(* IEC 61131-3 sources: volt/packages/volt-lsp-iec/libraries/Standard/3.5.18.0, 22 files *)

(* ---- CONCAT.pou ---- *)
FUNCTION CONCAT : STRING(255)
VAR_INPUT
	STR1 : STRING(255);
	STR2 : STRING(255);
END_VAR
VAR
	i : DINT;
	n : DINT;
END_VAR
(* STR2 after STR1, cut at the 255 the result holds *)
CONCAT := STR1;
n := UINT_TO_DINT(LEN_INTERNAL(STR1));
WHILE n + i < 255 AND STR2[i] <> 0 DO
	CONCAT[n + i] := STR2[i];
	i := i + 1;
END_WHILE
CONCAT[n + i] := 0;
END_FUNCTION

(* ---- DELETE.pou ---- *)
FUNCTION DELETE : STRING(255)
VAR_INPUT
	STR : STRING(255);
	LEN : INT;
	POS : INT;
END_VAR
VAR
	i : DINT;
	k : DINT;
	n : DINT;
	first : DINT;
	start : DINT;
	count : DINT;
END_VAR
(* LEN characters from POS, counting from 1. POSITION 0 IS NOT "DO NOTHING": the range starts at POS - 1, which may
   be negative, and what goes is the part of [POS - 1, POS - 1 + LEN) inside the string. DELETE('abcde', 2, 0) is
   'bcde' (measured str_delete_at_zero, 2026-09-19). *)
DELETE := STR;
IF LEN > 0 THEN
	n := UINT_TO_DINT(LEN_INTERNAL(STR));
	first := INT_TO_DINT(POS) - 1;
	start := MAX(first, 0);
	count := INT_TO_DINT(LEN) + MIN(first, 0);
	IF count > 0 AND start < n THEN
		k := start;
		FOR i := MIN(start + count, n) TO n - 1 DO
			DELETE[k] := STR[i];
			k := k + 1;
		END_FOR
		DELETE[k] := 0;
	END_IF
END_IF
END_FUNCTION

(* ---- FIND.pou ---- *)
FUNCTION FIND : INT
VAR_INPUT
	STR1 : STRING(255);
	STR2 : STRING(255);
END_VAR
VAR
	i : DINT;
	j : DINT;
	n1 : DINT;
	n2 : DINT;
END_VAR
(* where STR2 first starts in STR1, counting from 1; 0 when it does not occur, and FIND of '' is 0 *)
n1 := UINT_TO_DINT(LEN_INTERNAL(STR1));
n2 := UINT_TO_DINT(LEN_INTERNAL(STR2));
IF n2 > 0 THEN
	FOR i := 0 TO n1 - n2 DO
		j := 0;
		WHILE j < n2 AND STR1[i + j] = STR2[j] DO
			j := j + 1;
		END_WHILE
		IF j = n2 THEN
			FIND := DINT_TO_INT(i + 1);
			RETURN;
		END_IF
	END_FOR
END_IF
END_FUNCTION

(* ---- INSERT.pou ---- *)
FUNCTION INSERT : STRING(255)
VAR_INPUT
	STR1 : STRING(255);
	STR2 : STRING(255);
	POS : INT;
END_VAR
VAR
	i : DINT;
	k : DINT;
	n : DINT;
END_VAR
(* STR2 after the first POS characters of STR1. POS 0 prepends; a POS below 0 or past the end leaves STR1 as it was:
   INSERT('abc', 'XY', -1) is 'abc'. The result is cut at 255. *)
n := UINT_TO_DINT(LEN_INTERNAL(STR1));
IF POS < 0 OR POS > n THEN
	INSERT := STR1;
ELSE
	FOR i := 0 TO INT_TO_DINT(POS) - 1 DO
		INSERT[k] := STR1[i];
		k := k + 1;
	END_FOR
	i := 0;
	WHILE k < 255 AND STR2[i] <> 0 DO
		INSERT[k] := STR2[i];
		k := k + 1;
		i := i + 1;
	END_WHILE
	i := POS;
	WHILE k < 255 AND i < n DO
		INSERT[k] := STR1[i];
		k := k + 1;
		i := i + 1;
	END_WHILE
	INSERT[k] := 0;
END_IF
END_FUNCTION

(* ---- LEFT.pou ---- *)
FUNCTION LEFT : STRING(255)
VAR_INPUT
	STR : STRING(255);
	SIZE : INT;
END_VAR
VAR
	i : DINT;
	n : DINT;
END_VAR
(* SIZE clamps to the string: LEFT('abc', 5) is 'abc', LEFT('abc', -1) is '' *)
n := LIMIT(0, SIZE, UINT_TO_DINT(LEN_INTERNAL(STR)));
FOR i := 0 TO n - 1 DO
	LEFT[i] := STR[i];
END_FOR
LEFT[n] := 0;
END_FUNCTION

(* ---- LEN.pou ---- *)
FUNCTION LEN : INT
VAR_INPUT
	STR : STRING(255);
END_VAR
LEN := UINT_TO_INT(LEN_INTERNAL(STR));
END_FUNCTION

(* ---- LEN_INTERNAL.pou ---- *)
FUNCTION LEN_INTERNAL : UINT
VAR_IN_OUT
	STR : STRING(255);
END_VAR
(* the characters before the terminator: the one loop every other string function counts with *)
WHILE STR[LEN_INTERNAL] <> 0 DO
	LEN_INTERNAL := LEN_INTERNAL + 1;
END_WHILE
END_FUNCTION

(* ---- MEMCOPY_INTERNAL.pou ---- *)
FUNCTION MEMCOPY_INTERNAL : POINTER TO BYTE
VAR_INPUT
	PDEST : POINTER TO BYTE;
	PSRC : POINTER TO BYTE;
	DWSIZE : DWORD;
END_VAR
MEMCOPY_INTERNAL := PDEST;
WHILE DWSIZE > 0 DO
	PDEST^ := PSRC^;
	PDEST := PDEST + 1;
	PSRC := PSRC + 1;
	DWSIZE := DWSIZE - 1;
END_WHILE
END_FUNCTION

(* ---- MID.pou ---- *)
FUNCTION MID : STRING(255)
VAR_INPUT
	STR : STRING(255);
	LEN : INT;
	POS : INT;
END_VAR
VAR
	i : DINT;
	n : DINT;
	first : DINT;
	last : DINT;
END_VAR
(* POS counts from 1; a POS below 1 or a LEN at or below 0 selects nothing, and the span stops at the end *)
IF POS >= 1 AND LEN > 0 THEN
	n := UINT_TO_DINT(LEN_INTERNAL(STR));
	first := INT_TO_DINT(POS) - 1;
	last := first + INT_TO_DINT(LEN);
	i := first;
	WHILE i < n AND i < last DO
		MID[i - first] := STR[i];
		i := i + 1;
	END_WHILE
	MID[i - first] := 0;
END_IF
END_FUNCTION

(* ---- REPLACE.pou ---- *)
FUNCTION REPLACE : STRING(255)
VAR_INPUT
	STR1 : STRING(255);
	STR2 : STRING(255);
	L : INT;
	P : INT;
END_VAR
(* a DELETE, then an INSERT at P - 1 raised to 0. Every measured REPLACE agrees: REPLACE('abc', 'XY', 1, 0) is
   'XYabc' and REPLACE('abc', 'XY', 2, 5) is 'abc'. *)
REPLACE := INSERT(DELETE(STR1, L, P), STR2, MAX(P - 1, 0));
END_FUNCTION

(* ---- RIGHT.pou ---- *)
FUNCTION RIGHT : STRING(255)
VAR_INPUT
	STR : STRING(255);
	SIZE : INT;
END_VAR
VAR
	i : DINT;
	n : DINT;
	start : DINT;
END_VAR
n := UINT_TO_DINT(LEN_INTERNAL(STR));
start := n - LIMIT(0, SIZE, n);
FOR i := start TO n - 1 DO
	RIGHT[i - start] := STR[i];
END_FOR
RIGHT[n - start] := 0;
END_FUNCTION

(* ---- CTD.pou ---- *)
FUNCTION_BLOCK CTD
VAR_INPUT
	CD : BOOL;
	LOAD : BOOL;
	PV : WORD;
END_VAR
VAR_OUTPUT
	Q : BOOL;
	CV : WORD;
END_VAR
VAR
	M : BOOL;
END_VAR
IF LOAD THEN
	CV := PV;
ELSIF CD AND NOT M AND CV > 0 THEN
	CV := CV - 1;
END_IF
M := CD;
Q := CV = 0;
END_FUNCTION_BLOCK

(* ---- CTU.pou ---- *)
FUNCTION_BLOCK CTU
VAR_INPUT
	CU : BOOL;
	RESET : BOOL;
	PV : WORD;
END_VAR
VAR_OUTPUT
	Q : BOOL;
	CV : WORD;
END_VAR
VAR
	M : BOOL;
END_VAR
(* counts CU's rising edges, and stops at the top of the WORD rather than wrapping *)
IF RESET THEN
	CV := 0;
ELSIF CU AND NOT M AND CV < 16#FFFF THEN
	CV := CV + 1;
END_IF
M := CU;
Q := CV >= PV;
END_FUNCTION_BLOCK

(* ---- CTUD.pou ---- *)
FUNCTION_BLOCK CTUD
VAR_INPUT
	CU : BOOL;
	CD : BOOL;
	RESET : BOOL;
	LOAD : BOOL;
	PV : WORD;
END_VAR
VAR_OUTPUT
	QU : BOOL;
	QD : BOOL;
	CV : WORD;
END_VAR
VAR
	MU : BOOL;
	MD : BOOL;
	RU : BOOL;
	RD : BOOL;
END_VAR
(* RU and RD are the library's own variables, and this body has no use for them *)
IF RESET THEN
	CV := 0;
ELSIF LOAD THEN
	CV := PV;
ELSE
	IF CU AND NOT MU AND CV < 16#FFFF THEN
		CV := CV + 1;
	END_IF
	IF CD AND NOT MD AND CV > 0 THEN
		CV := CV - 1;
	END_IF
END_IF
MU := CU;
MD := CD;
QU := CV >= PV;
QD := CV = 0;
END_FUNCTION_BLOCK

(* ---- F_TRIG.pou ---- *)
FUNCTION_BLOCK F_TRIG
VAR_INPUT
	CLK : BOOL;
END_VAR
VAR_OUTPUT
	Q : BOOL;
END_VAR
VAR
	M : BOOL := TRUE;
END_VAR
(* M holds NOT CLK, which is why it starts TRUE: FALSE would report a falling edge on the first scan *)
Q := NOT CLK AND NOT M;
M := NOT CLK;
END_FUNCTION_BLOCK

(* ---- R_TRIG.pou ---- *)
FUNCTION_BLOCK R_TRIG
VAR_INPUT
	CLK : BOOL;
END_VAR
VAR_OUTPUT
	Q : BOOL;
END_VAR
VAR
	M : BOOL;
END_VAR
Q := CLK AND NOT M;
M := CLK;
END_FUNCTION_BLOCK

(* ---- RS.pou ---- *)
FUNCTION_BLOCK RS
VAR_INPUT
	SET : BOOL;
	RESET1 : BOOL;
END_VAR
VAR_OUTPUT
	Q1 : BOOL;
END_VAR
Q1 := NOT RESET1 AND (SET OR Q1);
END_FUNCTION_BLOCK

(* ---- RTC.pou ---- *)
FUNCTION_BLOCK RTC
VAR_INPUT
	EN : BOOL;
	PDT : DATE_AND_TIME;
END_VAR
VAR_OUTPUT
	Q : BOOL;
	CDT : DATE_AND_TIME;
END_VAR
VAR
	M : BOOL;
	DIFFTIME : TIME;
	LASTTIME : TIME := TIME#0ms;
	TIMEOFFSET : TIME := TIME#0ms;
	CURTIME : TIME;
END_VAR
(* CDT starts at PDT on EN's rising edge and runs with the clock; TIMEOFFSET carries the milliseconds a DT, which
   counts seconds, cannot hold yet *)
IF EN THEN
	CURTIME := TIME();
	IF NOT M THEN
		CDT := PDT;
		LASTTIME := CURTIME;
		TIMEOFFSET := TIME#0ms;
		M := TRUE;
	END_IF
	DIFFTIME := CURTIME - LASTTIME + TIMEOFFSET;
	CDT := DWORD_TO_DT(DT_TO_DWORD(CDT) + TIME_TO_DWORD(DIFFTIME) / 1000);
	TIMEOFFSET := DWORD_TO_TIME(TIME_TO_DWORD(DIFFTIME) MOD 1000);
	LASTTIME := CURTIME;
	Q := TRUE;
ELSE
	M := FALSE;
	Q := FALSE;
END_IF
END_FUNCTION_BLOCK

(* ---- SR.pou ---- *)
FUNCTION_BLOCK SR
VAR_INPUT
	SET1 : BOOL;
	RESET : BOOL;
END_VAR
VAR_OUTPUT
	Q1 : BOOL;
END_VAR
Q1 := SET1 OR (NOT RESET AND Q1);
END_FUNCTION_BLOCK

(* ---- TOF.pou ---- *)
FUNCTION_BLOCK TOF
VAR_INPUT
	IN : BOOL;
	PT : TIME;
END_VAR
VAR_OUTPUT
	Q : BOOL;
	ET : TIME;
END_VAR
VAR
	M : BOOL;
	STARTTIME : TIME;
END_VAR
(* Q follows IN up at once, and falls PT after IN has fallen *)
IF IN THEN
	Q := TRUE;
	ET := TIME#0ms;
	M := TRUE;
ELSE
	IF M THEN
		STARTTIME := TIME();
		M := FALSE;
	END_IF
	IF Q THEN
		ET := TIME() - STARTTIME;
		IF ET >= PT THEN
			Q := FALSE;
			ET := PT;
		END_IF
	END_IF
END_IF
END_FUNCTION_BLOCK

(* ---- TON.pou ---- *)
FUNCTION_BLOCK TON
VAR_INPUT
	IN : BOOL;
	PT : TIME;
END_VAR
VAR_OUTPUT
	Q : BOOL;
	ET : TIME;
END_VAR
VAR
	M : BOOL;
	STARTTIME : TIME;
END_VAR
(* Q rises once IN has been TRUE for PT; ET counts up to PT and holds there. TIME() is an operator of the language,
   not of this library: the one thing the library needs that ST cannot say by itself. *)
IF IN THEN
	IF NOT M THEN
		STARTTIME := TIME();
		M := TRUE;
	END_IF
	IF NOT Q THEN
		ET := TIME() - STARTTIME;
		IF ET >= PT THEN
			Q := TRUE;
			ET := PT;
		END_IF
	END_IF
ELSE
	Q := FALSE;
	ET := TIME#0ms;
	M := FALSE;
END_IF
END_FUNCTION_BLOCK

(* ---- TP.pou ---- *)
FUNCTION_BLOCK TP
VAR_INPUT
	IN : BOOL;
	PT : TIME;
END_VAR
VAR_OUTPUT
	Q : BOOL;
	ET : TIME;
END_VAR
VAR
	STARTTIME : TIME;
END_VAR
(* a pulse of PT on IN's rising edge, which IN falling does not cut short. Once no pulse runs and IN is FALSE,
   ET is 0 — in the very scan the pulse runs out, not the one after (recorded: lib_std_tp) — and ET = 0 is what arms
   the next pulse *)
IF Q THEN
	ET := TIME() - STARTTIME;
	IF ET >= PT THEN
		Q := FALSE;
		ET := PT;
	END_IF
ELSIF IN THEN
	IF ET = TIME#0ms THEN
		STARTTIME := TIME();
		Q := TRUE;
	END_IF
END_IF
IF NOT IN AND NOT Q THEN
	ET := TIME#0ms;
END_IF
END_FUNCTION_BLOCK
